// SIMATIC S7-200 project (STEP 7-Micro/WIN), CPU 224 CN REL 02.01

SYMBOL_TABLE USUARIO1
SB_1             I1.2     // Pulsador verde
SB_2             I1.3     // Pulsador rojo
QS               I1.4     // Emergencia
SA               I1.5     // Selector SA
PISTON_PEQ_ATR   I0.1     // Sensor magnetico de cilindro retraido
PISTON_PEQ_ADELANT I0.0     // Sensor magnetico de cilindro extendido
GRANDE_ADEL      I0.2     // Sensor magnetico de cilindro extendido
GRANDE_ATRAS     I0.3     // Sensor magnetico de cilindro retraido
presencia_superior I0.5     // S. fotoelectrico de presenscia en la parte superior del tubo
presencia_inferior I0.6     // S. fotoelectrico de presenscia en la parte inferior del tubo
posicion_final   I0.4     // S. pieza en posicion para la unidad de transporte
piston_peq       Q0.0     // Accionamiento cilindro neumatico superior
piston_grande    Q0.1     // Accionamiento cilindro neumatico inferior
HL1              Q0.7     // Señalizacion amarrilla
HL2              Q1.0     // Señalizacion verde
HL3              Q1.1     // Señalizacion roja
HL1_intermedio   M5.0
E0               M0.0     // Estado 0
E1               M0.1     // Estado 1
E2               M0.2     // Estado 2
E3               M0.3     // Estado 3
E4               M0.4     // Estado 4
E5               M0.5     // Estado 5
EM0              M0.6     // Estado de emergencia 0
EM1              M0.7     // Estado de emergencia 1
com_finalizado   V0.1     // Bit de comunicacion (hacia tranporte)
com_inicial      V0.0     // Bit de comunicacion (desde tranporte)
man_aut          M1.0     // Estado de manual y automatico
parada_momentanea M1.1     // Estado de la parada momentanea
END_SYMBOL_TABLE

ORGANIZATION_BLOCK PRINCIPAL:OB1
TITLE=PROGRAMA PRINCIPAL
BEGIN
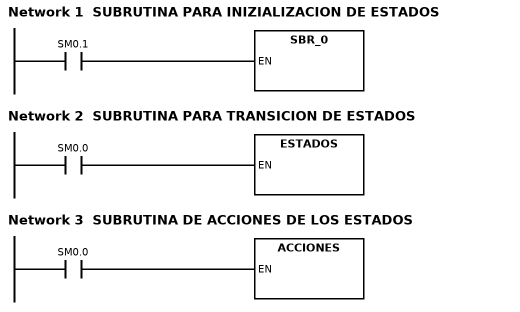
Network 1 // SUBRUTINA PARA INIZIALIZACION DE ESTADOS
LD     SM0.1
CALL   SBR_0:SBR0
Network 2 // SUBRUTINA PARA TRANSICION DE ESTADOS
LD     SM0.0
CALL   ESTADOS:SBR1
Network 3 // SUBRUTINA DE ACCIONES DE LOS ESTADOS
LD     SM0.0
CALL   ACCIONES:SBR2
END_ORGANIZATION_BLOCK

SUBROUTINE_BLOCK SBR_0:SBR0
TITLE=COMENTARIOS DE LA SUBRUTINA
BEGIN
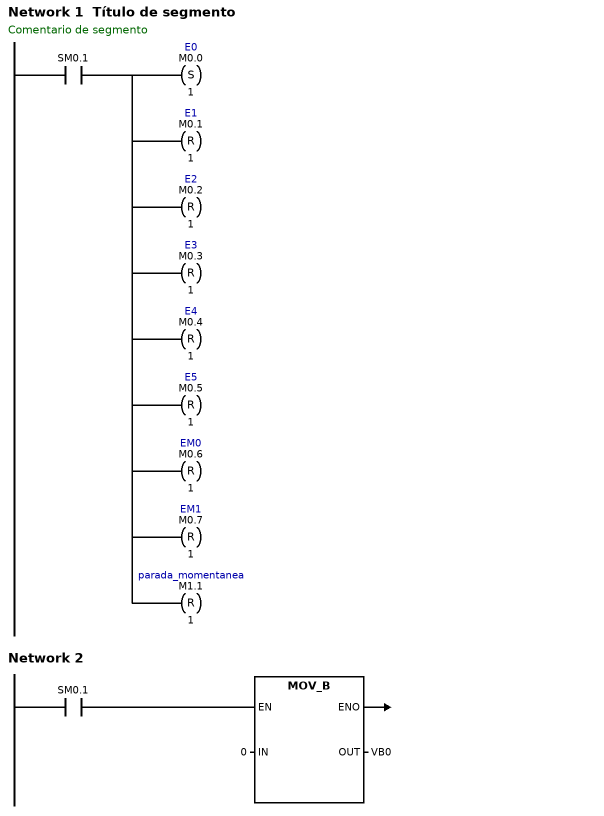
Network 1 // Título de segmento
// Comentario de segmento
LD     SM0.1
S      E0:M0.0, 1
R      E1:M0.1, 1
R      E2:M0.2, 1
R      E3:M0.3, 1
R      E4:M0.4, 1
R      E5:M0.5, 1
R      EM0:M0.6, 1
R      EM1:M0.7, 1
R      parada_momentanea:M1.1, 1
Network 2
LD     SM0.1
MOVB   0, VB0
END_SUBROUTINE_BLOCK

SUBROUTINE_BLOCK ESTADOS:SBR1
TITLE=TRANSICION DE ESTADOS
BEGIN
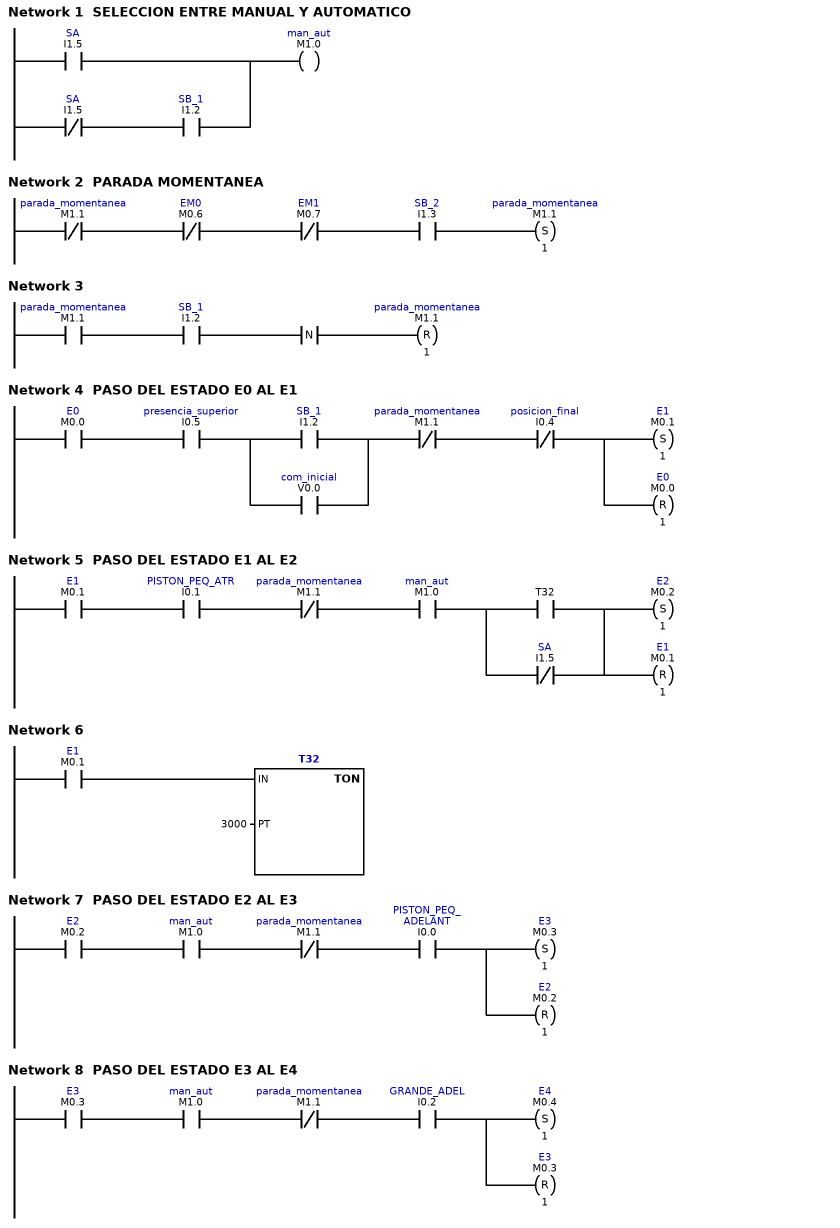
Network 1 // SELECCION ENTRE MANUAL Y AUTOMATICO
LD     SA:I1.5
LDN    SA:I1.5
A      SB_1:I1.2
OLD
=      man_aut:M1.0
Network 2 // PARADA MOMENTANEA
LDN    parada_momentanea:M1.1
AN     EM0:M0.6
AN     EM1:M0.7
A      SB_2:I1.3
S      parada_momentanea:M1.1, 1
Network 3
LD     parada_momentanea:M1.1
A      SB_1:I1.2
ED
R      parada_momentanea:M1.1, 1
Network 4 // PASO DEL ESTADO E0 AL E1
LD     E0:M0.0
A      presencia_superior:I0.5
LD     SB_1:I1.2
O      com_inicial:V0.0
ALD
AN     parada_momentanea:M1.1
AN     posicion_final:I0.4
S      E1:M0.1, 1
R      E0:M0.0, 1
Network 5 // PASO DEL ESTADO E1 AL E2
LD     E1:M0.1
A      PISTON_PEQ_ATR:I0.1
AN     parada_momentanea:M1.1
A      man_aut:M1.0
LD     T32
ON     SA:I1.5
ALD
S      E2:M0.2, 1
R      E1:M0.1, 1
Network 6
LD     E1:M0.1
TON    T32, 3000
Network 7 // PASO DEL ESTADO E2 AL E3
LD     E2:M0.2
A      man_aut:M1.0
AN     parada_momentanea:M1.1
A      PISTON_PEQ_ADELANT:I0.0
S      E3:M0.3, 1
R      E2:M0.2, 1
Network 8 // PASO DEL ESTADO E3 AL E4
LD     E3:M0.3
A      man_aut:M1.0
AN     parada_momentanea:M1.1
A      GRANDE_ADEL:I0.2
S      E4:M0.4, 1
R      E3:M0.3, 1
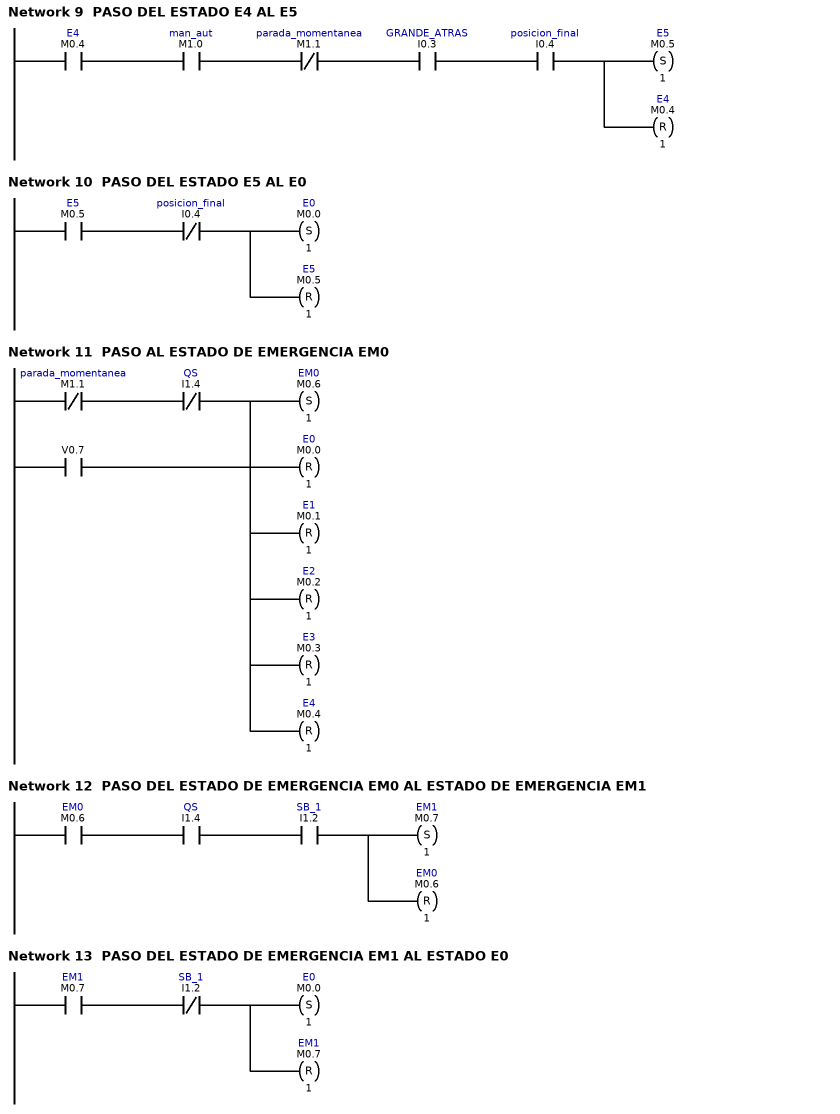
Network 9 // PASO DEL ESTADO E4 AL E5
LD     E4:M0.4
A      man_aut:M1.0
AN     parada_momentanea:M1.1
A      GRANDE_ATRAS:I0.3
A      posicion_final:I0.4
S      E5:M0.5, 1
R      E4:M0.4, 1
Network 10 // PASO DEL ESTADO E5 AL E0
LD     E5:M0.5
AN     posicion_final:I0.4
S      E0:M0.0, 1
R      E5:M0.5, 1
Network 11 // PASO AL ESTADO DE EMERGENCIA EM0
LDN    parada_momentanea:M1.1
AN     QS:I1.4
O      V0.7
S      EM0:M0.6, 1
R      E0:M0.0, 1
R      E1:M0.1, 1
R      E2:M0.2, 1
R      E3:M0.3, 1
R      E4:M0.4, 1
Network 12 // PASO DEL ESTADO DE EMERGENCIA EM0 AL ESTADO DE EMERGENCIA EM1
LD     EM0:M0.6
A      QS:I1.4
A      SB_1:I1.2
S      EM1:M0.7, 1
R      EM0:M0.6, 1
Network 13 // PASO DEL ESTADO DE EMERGENCIA EM1 AL ESTADO E0
LD     EM1:M0.7
AN     SB_1:I1.2
S      E0:M0.0, 1
R      EM1:M0.7, 1
END_SUBROUTINE_BLOCK

SUBROUTINE_BLOCK ACCIONES:SBR2
TITLE=ACCIONES EN ESTADOS
BEGIN
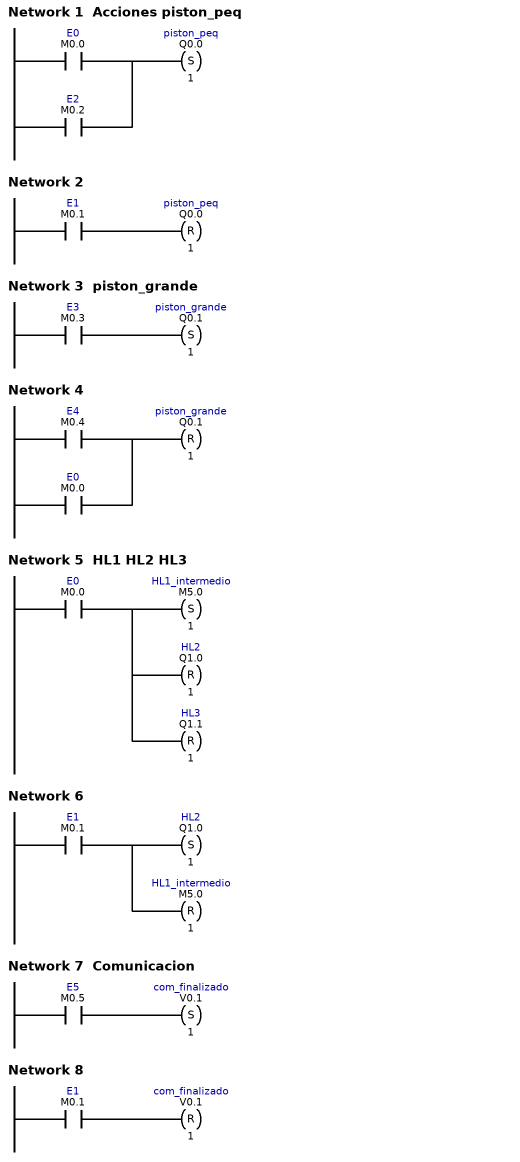
Network 1 // Acciones
piston_peq
LD     E0:M0.0
O      E2:M0.2
S      piston_peq:Q0.0, 1
Network 2
LD     E1:M0.1
R      piston_peq:Q0.0, 1
Network 3 // piston_grande
LD     E3:M0.3
S      piston_grande:Q0.1, 1
Network 4
LD     E4:M0.4
O      E0:M0.0
R      piston_grande:Q0.1, 1
Network 5 // HL1
HL2
HL3
LD     E0:M0.0
S      HL1_intermedio:M5.0, 1
R      HL2:Q1.0, 1
R      HL3:Q1.1, 1
Network 6
LD     E1:M0.1
S      HL2:Q1.0, 1
R      HL1_intermedio:M5.0, 1
Network 7 // Comunicacion
LD     E5:M0.5
S      com_finalizado:V0.1, 1
Network 8
LD     E1:M0.1
R      com_finalizado:V0.1, 1
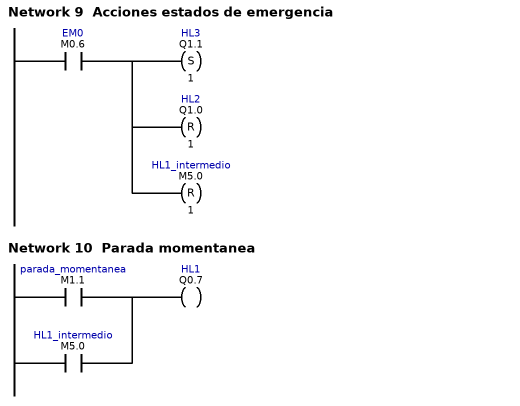
Network 9 // Acciones estados de emergencia
LD     EM0:M0.6
S      HL3:Q1.1, 1
R      HL2:Q1.0, 1
R      HL1_intermedio:M5.0, 1
Network 10 // Parada momentanea
LD     parada_momentanea:M1.1
O      HL1_intermedio:M5.0
=      HL1:Q0.7
END_SUBROUTINE_BLOCK
